(* PLC project PR_HIPOTTestSeq_Soft2.0 1_workflow_cd2a65_PLC, SiemensToBackhoff Siemens TIA Portal → Beckhoff TwinCAT PLCopen Converter 2.2 *)
(* stored: creationDateTime 2026-10-12T09:24:44.936111, modificationDateTime 2026-10-12T09:24:44.936111 *)

FUNCTION_BLOCK PR_HIPOTTestSeq_Soft2.0 1_workflow_cd2a65
VAR_INPUT
	iAutoRunning : BOOL;
	iFaultReset : BOOL;
	iHiPotProbeUp : BOOL;
	iHiPotTestOver : BOOL;
	iHiPotTestProbeDown : BOOL;
	iPartPresent : BOOL;
	iPressProbeUp : BOOL;
	iReset_fault : BOOL;
	iShuttleAtHiPotTest : BOOL;
	iSstMode : BOOL;
	iSstPB : BOOL;
	iStartFrmShuttleSeq : BOOL;
	iTestProbeDown : BOOL;
	iTestProbeUp : BOOL;
	iTestProbesUp : BOOL;
	iThicknessTestOver : BOOL;
	iScanOK : BOOL;
	iScanNOK : BOOL;
	iRetryCount : INT;
	iForcedAccept : BOOL;
	iRetry : BOOL;
END_VAR
VAR_OUTPUT
	qHiPotTestOver : BOOL;
	qStateNo : INT;
	qMessage : ARRAY[0..2] OF BOOL;
END_VAR
VAR
	c20_ChkRecoveryStatus_T1 : BOOL;
	c20_ChkRecoveryStatus_T2 : BOOL;
	c20_ChkRecoveryStatus_T3 : BOOL;
	c20_ChkRecoveryStatus_T4 : BOOL;
	c50_ChkPartPresentShuttlePos_T1 : BOOL;
	c50_ChkPartPresentShuttlePos_T2 : BOOL;
	s100_WtHiPotTestProbesDown : BOOL;
	s100_WtHiPotTestProbesDown_T1 : BOOL;
	s10_WtStartFrmShuttleSeq : BOOL;
	s10_WtStartFrmShuttleSeq_T1 : BOOL;
	s110_WtHiPotTestOver : BOOL;
	s110_WtHiPotTestOver_T1 : BOOL;
	s120_WtHiPotProbeUp : BOOL;
	s120_WtHiPotProbeUp_T1 : BOOL;
	s130_WtPressProbesUp : BOOL;
	s130_WtPressProbesUp_T1 : BOOL;
	s140_WtStartLow : BOOL;
	s140_WtStartLow_T1 : BOOL;
	s1_WtResetRel : BOOL;
	s1_WtResetRel_T1 : BOOL;
	s20_ChkRecoveryStatus : BOOL;
	s20_ChkRecoveryStatus_T1 : BOOL;
	s20_ChkRecoveryStatus_T2 : BOOL;
	s20_ChkRecoveryStatus_T3 : BOOL;
	s20_ChkRecoveryStatus_T4 : BOOL;
	s30_WtOperatorAck : BOOL;
	s30_WtOperatorAck_T1 : BOOL;
	s40_WtAllSlidesHome : BOOL;
	s40_WtAllSlidesHome_T1 : BOOL;
	s50_ChkPartPresentShuttlePos : BOOL;
	s50_ChkPartPresentShuttlePos_T1 : BOOL;
	s50_ChkPartPresentShuttlePos_T2 : BOOL;
	s75_WtScanOver : BOOL;
	s75_WtScanOver_T1 : BOOL;
	s75_WtScanOver_T2 : BOOL;
	s76_ChkReryCountOver : BOOL;
	s76_ChkRetryCountOver_T1 : BOOL;
	s76_ChkRetryCountOver_T2 : BOOL;
	s77_WtOperatorDecision : BOOL;
	s77_WtOperatorDecision_T1 : BOOL;
	s77_WtOperatorDecision_T2 : BOOL;
	s70_WtPartPresentShuttlePos : BOOL;
	s70_WtPartPresentShuttlePos_T1 : BOOL;
	s80_WtTestProbeDown : BOOL;
	s80_WtTestProbeDown_T1 : BOOL;
	s90_WtThicknessTestOver : BOOL;
	s90_WtThicknessTestOver_T1 : BOOL;
	sAbnormalStatus : BOOL;
	sHiPotTestInProgress : BOOL;
	sSst : BOOL;
	sSstPulse : BOOL;
	sSstRise : R_TRIG;
	sStWtResetRel : BOOL;
	sStWtResetRel_T1 : BOOL;
	sThicknessTestInProgress : BOOL;
	sScanRetryCount : INT;
END_VAR
VAR_TEMP
	tOne : BOOL;
END_VAR
  VAR  (* added by the conversion: wires and edge detectors of the diagram *)
    _w24 : BOOL;
    _w26 : BOOL;
    _w39 : BOOL;
    _w41 : BOOL;
    _w42 : BOOL;
    _w55 : BOOL;
    _w58 : BOOL;
    _w59 : BOOL;
    _w102 : BOOL;
    _w105 : BOOL;
    _w106 : BOOL;
    _w107 : BOOL;
    _w108 : BOOL;
    _w109 : BOOL;
    _w122 : BOOL;
    _w124 : BOOL;
    _w125 : BOOL;
    _w139 : BOOL;
    _w141 : BOOL;
    _w142 : BOOL;
    _w178 : BOOL;
    _w180 : BOOL;
    _w181 : BOOL;
    _w182 : BOOL;
    _w200 : BOOL;
    _w202 : BOOL;
    _w203 : BOOL;
    _w219 : BOOL;
    _w223 : BOOL;
    _w224 : BOOL;
    _w225 : BOOL;
    _GT237_ENO : BOOL;
    _GT237_OUT : BOOL;
    _LE241_ENO : BOOL;
    _LE241_OUT : BOOL;
    _w245 : BOOL;
    _w247 : BOOL;
    _w248 : BOOL;
    _w249 : BOOL;
    _w265 : BOOL;
    _w267 : BOOL;
    _w268 : BOOL;
    _w269 : BOOL;
    _w282 : BOOL;
    _w286 : BOOL;
    _w287 : BOOL;
    _w300 : BOOL;
    _w303 : BOOL;
    _w304 : BOOL;
    _w321 : BOOL;
    _w323 : BOOL;
    _w324 : BOOL;
    _w337 : BOOL;
    _w340 : BOOL;
    _w341 : BOOL;
    _w358 : BOOL;
    _w360 : BOOL;
    _w361 : BOOL;
    _w374 : BOOL;
    _w376 : BOOL;
    _w377 : BOOL;
    _w390 : BOOL;
    _w392 : BOOL;
    _w393 : BOOL;
  END_VAR

(* LD diagram, written out as Structured Text *)
(* Network 1 *)
(* Create Single Step Pulse bit *)
(* Create Single Step bit *)
(* Transition for STATE Num:0 Reset Released *)
(* STATE Num:0 Reset Released *)
(* Transition for STATE Num:1 WtResetRel *)
(* STATE Num:1 WtResetRel *)
(* Transition for STATE Num:10 WtStartFrmShuttleSeq *)
(* STATE Num:10 WtStartFrmShuttleSeq *)
(* Condition1 for STATE Num:20 ChkRecoveryStatus *)
(* Condition2 for STATE Num:20 ChkRecoveryStatus *)
(* Condition3 for STATE Num:20 ChkRecoveryStatus *)
(* Condition4 for STATE Num:20 ChkRecoveryStatus *)
(* Transition for STATE Num:20 ChkRecoveryStatus *)
(* STATE Num:20 ChkRecoveryStatus *)
(* Transition for STATE Num:30 WtOperatorAck *)
(* STATE Num:30 WtOperatorAck *)
(* Transition for STATE Num:40 WtAllSlidesHome *)
(* STATE Num:40 WtAllSlidesHome *)
(* Actions for STATE Num:40 WtAllSlidesHome - qMessage[1] if TestProbe not up *)
(* Actions for STATE Num:40 WtAllSlidesHome - qMessage[2] if PressProbe not up *)
(* Condition1 for STATE Num:50 ChkPartPresentShuttlePos *)
(* Condition2 for STATE Num:50 ChkPartPresentShuttlePos *)
(* Transition for STATE Num:50 ChkPartPresentShuttlePos *)
(* STATE Num:50 ChkPartPresentShuttlePos *)
(* Actions for STATE Num:50 ChkPartPresentShuttlePos *)
(* Transition for STATE Num:70 WtPartPresentShuttlePos *)
(* STATE Num:70 WtPartPresentShuttlePos *)
(* Transition for STATE Num:75 WtScan Over *)
(* STATE Num:75 WtScanOver *)
(* Transition for STATE Num:76 CheckRetryCountOver *)
(* STATE Num:76 CheckRetryCount *)
(* Transition for STATE Num:77 wair for operator Decision *)
(* STATE Num:77 wait For Operator Decision *)
(* Transition for STATE Num:80 WtTestProbeDown *)
(* STATE Num:80 WtTestProbeDown *)
(* Transition for STATE Num:90 WtThicknessTestOver *)
(* STATE Num:90 WtThicknessTestOver *)
(* Actions for STATE Num:90 WtThicknessTestOver *)
(* Transition for STATE Num:100 WtHiPotTestProbesDown *)
(* STATE Num:100 WtHiPotTestProbesDown *)
(* Transition for STATE Num:110 WtHiPotTestOver *)
(* STATE Num:110 WtHiPotTestOver *)
(* Actions for STATE Num:110 WtHiPotTestOver *)
(* Transition for STATE Num:120 WtHiPotProbeUp *)
(* STATE Num:120 WtHiPotProbeUp *)
(* Transition for STATE Num:130 WtPressProbesUp *)
(* STATE Num:130 WtPressProbesUp *)
(* Transition for STATE Num:140 WtStartLow *)
(* STATE Num:140 WtStartLow *)
(* Actions for STATE Num:140 WtStartLow - qHiPotTestOver *)
(* Actions for STATE Num:140 WtStartLow - Reset sHiPotTestInProgress on transition *)
(* Actions for STATE Num:140 WtStartLow - Reset sThicknessTestInProgress on transition *)
tOne := tOne OR NOT tOne;
sSstRise(CLK := iSstPB);
sSstPulse := sSstRise.Q;
sSst := iSstMode AND sSstPulse OR NOT iSstMode;
sStWtResetRel_T1 := sStWtResetRel AND iAutoRunning;
_w24 := sStWtResetRel;
_w26 := (_w24 OR NOT iAutoRunning) AND NOT sStWtResetRel_T1;
sStWtResetRel := _w26;
IF _w26 THEN qStateNo := 0; END_IF;
s1_WtResetRel_T1 := s1_WtResetRel AND NOT sStWtResetRel AND sSst AND iAutoRunning;
_w39 := s1_WtResetRel;
_w41 := (_w39 OR sStWtResetRel_T1) AND NOT sStWtResetRel;
_w42 := _w41 AND NOT s1_WtResetRel_T1;
s1_WtResetRel := _w42;
IF _w42 THEN qStateNo := 1; END_IF;
s10_WtStartFrmShuttleSeq_T1 := s10_WtStartFrmShuttleSeq AND NOT sStWtResetRel AND sSst AND iStartFrmShuttleSeq;
_w55 := s10_WtStartFrmShuttleSeq;
_w58 := (_w55 OR s1_WtResetRel_T1 OR s140_WtStartLow_T1) AND NOT sStWtResetRel;
_w59 := _w58 AND NOT s10_WtStartFrmShuttleSeq_T1;
s10_WtStartFrmShuttleSeq := _w59;
IF _w59 THEN qStateNo := 10; END_IF;
c20_ChkRecoveryStatus_T1 := sAbnormalStatus;
c20_ChkRecoveryStatus_T2 := sHiPotTestInProgress;
c20_ChkRecoveryStatus_T3 := sThicknessTestInProgress;
c20_ChkRecoveryStatus_T4 := NOT sAbnormalStatus AND NOT sHiPotTestInProgress AND NOT sThicknessTestInProgress;
s20_ChkRecoveryStatus_T1 := s20_ChkRecoveryStatus AND NOT sStWtResetRel AND sSst AND c20_ChkRecoveryStatus_T1;
s20_ChkRecoveryStatus_T2 := s20_ChkRecoveryStatus AND NOT sStWtResetRel AND sSst AND NOT s20_ChkRecoveryStatus_T1 AND c20_ChkRecoveryStatus_T2;
s20_ChkRecoveryStatus_T3 := s20_ChkRecoveryStatus AND NOT sStWtResetRel AND sSst AND NOT s20_ChkRecoveryStatus_T1 AND NOT s20_ChkRecoveryStatus_T1 AND NOT s20_ChkRecoveryStatus_T2 AND c20_ChkRecoveryStatus_T3;
s20_ChkRecoveryStatus_T4 := s20_ChkRecoveryStatus AND NOT sStWtResetRel AND sSst AND NOT s20_ChkRecoveryStatus_T1 AND NOT s20_ChkRecoveryStatus_T1 AND NOT s20_ChkRecoveryStatus_T2 AND NOT s20_ChkRecoveryStatus_T1 AND NOT s20_ChkRecoveryStatus_T2 AND NOT s20_ChkRecoveryStatus_T3 AND c20_ChkRecoveryStatus_T4;
_w102 := s20_ChkRecoveryStatus;
_w105 := (_w102 OR s10_WtStartFrmShuttleSeq_T1 OR s30_WtOperatorAck_T1) AND NOT sStWtResetRel;
_w106 := _w105 AND NOT s20_ChkRecoveryStatus_T1;
_w107 := _w106 AND NOT s20_ChkRecoveryStatus_T2;
_w108 := _w107 AND NOT s20_ChkRecoveryStatus_T3;
_w109 := _w108 AND NOT s20_ChkRecoveryStatus_T4;
s20_ChkRecoveryStatus := _w109;
IF _w109 THEN qStateNo := 20; END_IF;
s30_WtOperatorAck_T1 := s30_WtOperatorAck AND NOT sStWtResetRel AND sSst AND iFaultReset;
_w122 := s30_WtOperatorAck;
_w124 := (_w122 OR s20_ChkRecoveryStatus_T1) AND NOT sStWtResetRel;
_w125 := _w124 AND NOT s30_WtOperatorAck_T1;
s30_WtOperatorAck := _w125;
IF _w125 THEN qStateNo := 30; END_IF;
s40_WtAllSlidesHome_T1 := s40_WtAllSlidesHome AND NOT sStWtResetRel AND sSst AND iTestProbeUp AND iPressProbeUp;
_w139 := s40_WtAllSlidesHome;
_w141 := (_w139 OR s20_ChkRecoveryStatus_T4) AND NOT sStWtResetRel;
_w142 := _w141 AND NOT s40_WtAllSlidesHome_T1;
s40_WtAllSlidesHome := _w142;
IF _w142 THEN qStateNo := 40; END_IF;
qMessage[1] := s40_WtAllSlidesHome AND NOT iTestProbeUp;
qMessage[2] := s40_WtAllSlidesHome AND NOT iPressProbeUp;
c50_ChkPartPresentShuttlePos_T1 := NOT iPartPresent OR NOT iShuttleAtHiPotTest;
c50_ChkPartPresentShuttlePos_T2 := iPartPresent AND iShuttleAtHiPotTest;
s50_ChkPartPresentShuttlePos_T1 := s50_ChkPartPresentShuttlePos AND NOT sStWtResetRel AND sSst AND c50_ChkPartPresentShuttlePos_T1;
s50_ChkPartPresentShuttlePos_T2 := s50_ChkPartPresentShuttlePos AND NOT sStWtResetRel AND sSst AND NOT s50_ChkPartPresentShuttlePos_T1 AND c50_ChkPartPresentShuttlePos_T2;
_w178 := s50_ChkPartPresentShuttlePos;
_w180 := (_w178 OR s40_WtAllSlidesHome_T1) AND NOT sStWtResetRel;
_w181 := _w180 AND NOT s50_ChkPartPresentShuttlePos_T1;
_w182 := _w181 AND NOT s50_ChkPartPresentShuttlePos_T2;
s50_ChkPartPresentShuttlePos := _w182;
IF _w182 THEN qStateNo := 50; END_IF;
qMessage[0] := s50_ChkPartPresentShuttlePos;
s70_WtPartPresentShuttlePos_T1 := s70_WtPartPresentShuttlePos AND NOT sStWtResetRel AND sSst AND iPartPresent AND iShuttleAtHiPotTest;
_w200 := s70_WtPartPresentShuttlePos;
_w202 := (_w200 OR s50_ChkPartPresentShuttlePos_T1) AND NOT sStWtResetRel;
_w203 := _w202 AND NOT s70_WtPartPresentShuttlePos_T1;
s70_WtPartPresentShuttlePos := _w203;
IF _w203 THEN qStateNo := 70; END_IF;
s75_WtScanOver_T1 := s75_WtScanOver AND NOT sStWtResetRel AND sSst AND iScanNOK;
s75_WtScanOver_T2 := s75_WtScanOver AND NOT sStWtResetRel AND sSst AND NOT s75_WtScanOver_T1 AND iScanOK;
_w219 := s75_WtScanOver;
_w223 := (_w219 OR s70_WtPartPresentShuttlePos_T1 OR s76_ChkRetryCountOver_T2 OR s77_WtOperatorDecision_T2) AND NOT sStWtResetRel;
_w224 := _w223 AND NOT s75_WtScanOver_T1;
_w225 := _w224 AND NOT s75_WtScanOver_T2;
s75_WtScanOver := _w225;
IF _w225 THEN qStateNo := 75; END_IF;
_GT237_OUT := GT(EN := s76_ChkReryCountOver AND NOT sStWtResetRel AND sSst, IN1 := sScanRetryCount, IN2 := iRetryCount, ENO => _GT237_ENO);
s76_ChkRetryCountOver_T1 := _GT237_OUT;
_LE241_OUT := LE(EN := s76_ChkReryCountOver AND NOT sStWtResetRel AND sSst AND NOT s76_ChkRetryCountOver_T1, IN1 := sScanRetryCount, IN2 := iRetryCount, ENO => _LE241_ENO);
s76_ChkRetryCountOver_T2 := _LE241_OUT;
_w245 := s76_ChkReryCountOver;
_w247 := (_w245 OR s75_WtScanOver_T1) AND NOT sStWtResetRel;
_w248 := _w247 AND NOT s76_ChkRetryCountOver_T1;
_w249 := _w248 AND NOT s76_ChkRetryCountOver_T2;
s76_ChkReryCountOver := _w249;
IF _w249 THEN qStateNo := 76; END_IF;
s77_WtOperatorDecision_T1 := s77_WtOperatorDecision AND NOT sStWtResetRel AND sSst AND iForcedAccept;
s77_WtOperatorDecision_T2 := s77_WtOperatorDecision AND NOT sStWtResetRel AND sSst AND NOT s77_WtOperatorDecision_T1 AND iRetry;
_w265 := s77_WtOperatorDecision;
_w267 := (_w265 OR s76_ChkRetryCountOver_T1) AND NOT sStWtResetRel;
_w268 := _w267 AND NOT s77_WtOperatorDecision_T1;
_w269 := _w268 AND NOT s77_WtOperatorDecision_T2;
s77_WtOperatorDecision := _w269;
IF _w269 THEN qStateNo := 77; END_IF;
s80_WtTestProbeDown_T1 := s80_WtTestProbeDown AND NOT sStWtResetRel AND sSst AND iTestProbeDown;
_w282 := s80_WtTestProbeDown;
_w286 := (_w282 OR s75_WtScanOver_T2 OR s50_ChkPartPresentShuttlePos_T2 OR s77_WtOperatorDecision_T1) AND NOT sStWtResetRel;
_w287 := _w286 AND NOT s80_WtTestProbeDown_T1;
s80_WtTestProbeDown := _w287;
IF _w287 THEN qStateNo := 80; END_IF;
s90_WtThicknessTestOver_T1 := s90_WtThicknessTestOver AND NOT sStWtResetRel AND sSst AND iThicknessTestOver;
_w300 := s90_WtThicknessTestOver;
_w303 := (_w300 OR s80_WtTestProbeDown_T1 OR s20_ChkRecoveryStatus_T3) AND NOT sStWtResetRel;
_w304 := _w303 AND NOT s90_WtThicknessTestOver_T1;
s90_WtThicknessTestOver := _w304;
IF _w304 THEN qStateNo := 90; END_IF;
sThicknessTestInProgress := s90_WtThicknessTestOver;
s100_WtHiPotTestProbesDown_T1 := s100_WtHiPotTestProbesDown AND NOT sStWtResetRel AND sSst AND iHiPotTestProbeDown;
_w321 := s100_WtHiPotTestProbesDown;
_w323 := (_w321 OR s90_WtThicknessTestOver_T1) AND NOT sStWtResetRel;
_w324 := _w323 AND NOT s100_WtHiPotTestProbesDown_T1;
s100_WtHiPotTestProbesDown := _w324;
IF _w324 THEN qStateNo := 100; END_IF;
s110_WtHiPotTestOver_T1 := s110_WtHiPotTestOver AND NOT sStWtResetRel AND sSst AND iHiPotTestOver;
_w337 := s110_WtHiPotTestOver;
_w340 := (_w337 OR s100_WtHiPotTestProbesDown_T1 OR s20_ChkRecoveryStatus_T2) AND NOT sStWtResetRel;
_w341 := _w340 AND NOT s110_WtHiPotTestOver_T1;
s110_WtHiPotTestOver := _w341;
IF _w341 THEN qStateNo := 110; END_IF;
sHiPotTestInProgress := s110_WtHiPotTestOver;
s120_WtHiPotProbeUp_T1 := s120_WtHiPotProbeUp AND NOT sStWtResetRel AND sSst AND iHiPotProbeUp;
_w358 := s120_WtHiPotProbeUp;
_w360 := (_w358 OR s110_WtHiPotTestOver_T1) AND NOT sStWtResetRel;
_w361 := _w360 AND NOT s120_WtHiPotProbeUp_T1;
s120_WtHiPotProbeUp := _w361;
IF _w361 THEN qStateNo := 120; END_IF;
s130_WtPressProbesUp_T1 := s130_WtPressProbesUp AND NOT sStWtResetRel AND sSst AND iTestProbesUp;
_w374 := s130_WtPressProbesUp;
_w376 := (_w374 OR s120_WtHiPotProbeUp_T1) AND NOT sStWtResetRel;
_w377 := _w376 AND NOT s130_WtPressProbesUp_T1;
s130_WtPressProbesUp := _w377;
IF _w377 THEN qStateNo := 130; END_IF;
s140_WtStartLow_T1 := s140_WtStartLow AND NOT sStWtResetRel AND sSst AND NOT iStartFrmShuttleSeq;
_w390 := s140_WtStartLow;
_w392 := (_w390 OR s130_WtPressProbesUp_T1) AND NOT sStWtResetRel;
_w393 := _w392 AND NOT s140_WtStartLow_T1;
s140_WtStartLow := _w393;
IF _w393 THEN qStateNo := 140; END_IF;
qHiPotTestOver := s140_WtStartLow;
sHiPotTestInProgress := s140_WtStartLow AND NOT iStartFrmShuttleSeq;
sThicknessTestInProgress := s140_WtStartLow AND NOT iStartFrmShuttleSeq;
END_FUNCTION_BLOCK
